// Pilote du système planaire (docs/05 § 6). Le séquenceur ne donne que des destinations ; trajets et évitement
// de collision sont faits par le système planaire. FB_PlanarSim l'implémente en simulation ; le pilote Tc3 Planar
// (projet de la machine ou bibliothèque à venir) implémente la même interface.
INTERFACE I_PlanarDriver

METHOD Activate : BOOL              // TRUE quand le système est actif
VAR_INPUT
    bEnable : BOOL;
END_VAR
END_METHOD

METHOD MoveTo : BOOL                // TRUE si la commande est acceptée
VAR_INPUT
    nMover : USINT;
    stPos : ST_Position;
    fVelocity : LREAL;               // mm/s, override déjà appliqué par le pilote
    fAcceleration : LREAL;
END_VAR
END_METHOD

METHOD StopAll
END_METHOD

METHOD StopMover                    // arrêt contrôlé d'un mover (mode manuel)
VAR_INPUT
    nMover : USINT;
END_VAR
END_METHOD

METHOD AckError
END_METHOD

METHOD Cycle
VAR_INPUT
    fOverride : LREAL;               // override machine effectif, %
END_VAR
END_METHOD

METHOD MoverPosition : ST_Position
VAR_INPUT
    nMover : USINT;
END_VAR
END_METHOD

METHOD MoverMoving : BOOL
VAR_INPUT
    nMover : USINT;
END_VAR
END_METHOD

METHOD MoverDetected : BOOL
VAR_INPUT
    nMover : USINT;
END_VAR
END_METHOD

METHOD SetInitialPosition           // simulation : poser un mover sur le plan
VAR_INPUT
    nMover : USINT;
    stPos : ST_Position;
END_VAR
END_METHOD

PROPERTY Active : BOOL
GET
END_GET
END_PROPERTY

PROPERTY ErrorCode : UINT          // 0 ou erreur du type Système planaire (100 collision, 101 mover non détecté, 102 groupe)
GET
END_GET
END_PROPERTY

PROPERTY ErrorSubCode : UDINT
GET
END_GET
END_PROPERTY

END_INTERFACE

(* stored: Version 1.1.0.1, ProductVersion 3.1.4024.12
   Itf I_PlanarDriver: Id {e8f3f56c-07c1-5291-a0a2-fe146669344b}
   Method Activate: Id {72cfe9e8-c075-5cf8-9006-3301ccef908f}
   Method MoveTo: Id {7c93dbc3-2513-50c9-bcfe-e11b12e9e05f}
   Method StopAll: Id {de5b2d4c-a564-5d9a-b000-091f2981a608}
   Method StopMover: Id {805f4b8f-c407-58aa-8384-9de63a2828df}
   Method AckError: Id {91f973cb-223b-5e54-b3f4-a610e2754a14}
   Method Cycle: Id {7b9a37ad-85c9-52b5-8267-62ee424383dc}
   Method MoverPosition: Id {07c6bfb1-66f2-578c-87a1-5dff44ba935e}
   Method MoverMoving: Id {2b504c70-e2d8-56a4-9b0b-e6dd951ed423}
   Method MoverDetected: Id {e58b222a-fcde-54cc-a9b2-a16b791359fd}
   Method SetInitialPosition: Id {1bac688d-1867-5144-848c-c6322576c1c2}
   Property Active: Id {c67b5b2d-99b7-52c4-b0b0-240e555bbee4}
   Get Get: Id {c94b79a9-f3d2-50e3-bb82-6b6b6e9cff0f}
   Property ErrorCode: Id {7c85e702-7293-534f-b278-9b2f43d33299}
   Get Get: Id {2ca6d252-8f88-5cd8-b10c-a98d41e5f2b4}
   Property ErrorSubCode: Id {0d533be9-d15d-5c80-8499-333993b548d3}
   Get Get: Id {bf5f51b5-d3e5-5b7c-a3bd-b24f6e833f28} *)
